(* IEC 61131-3 sources: repolevel_ST_code_completion/dataset/project_code/four-level_elevator_control/global, 3 files *)

(* ---- GVL_Input.st ---- *)
VAR_GLOBAL
	IGoFloor	:	ARRAY[1..MaxNumFloor] OF BOOL;  //电梯里面
	ICallHelp	:	BOOL;
	IClose		:	BOOL;
	IOpen		:	BOOL;
	IIsClose	:	BOOL;
	IIsOpen		:	BOOL;

	IIsFloor	:	ARRAY[1..MaxNumFloor] OF BOOL := [TRUE];//电梯停在一层

	IFloorUp	:	ARRAY[1..MaxNumFloor - 1] OF BOOL; //电梯外面
	IFloorDown	:	ARRAY[2..MaxNumFloor] OF BOOL;

	IReset		:	BOOL;
	IRespondHelp	:	BOOL;
END_VAR

(* ---- GVL_Memory.st ---- *)
VAR_GLOBAL CONSTANT
	MaxNumFloor	:	USINT := 4;
END_VAR
VAR_GLOBAL
	Tar_Dir	:	Target_Direction;
END_VAR

(* ---- GVL_Output.st ---- *)
VAR_GLOBAL
	QMotorPositiveRun	:	BOOL;    //电梯处于向上运动状态
	QMotorNegativeRun	:	BOOL; //电梯处于向下运动状态
	QClose	:	BOOL := TRUE;    //电梯是处于关闭状态
	QOpen	:	BOOL;               //电梯是处于打开状态
	QHelpBeer	:	BOOL;        //报警灯是亮还是灭

	QGoFloorLed	:	ARRAY[1..MaxNumFloor] OF BOOL;   //电梯内“1/2/3/4”按钮，为TRUE时，按钮亮

	QFloorUpLed	:	ARRAY[1..MaxNumFloor - 1] OF BOOL;   //楼层中3个“上”按钮，为TRUE时，按钮亮
	QFloorDownLed	:	ARRAY[2..MaxNumFloor] OF BOOL;   //楼层中3个“下”按钮，为TRUE时，按钮亮
END_VAR
